Fanuc KAREL source: compact_preamble.KL

PROGRAM KB00046
%NOLOCKGROUP
%ENVIRONMENT FDEV
VAR
P1 : STRING[80];P2 : STRING[80];P3:BOOLEAN;P4:BOOLEAN;P5:INTEGER
BEGIN
P1='A'
P2='A'
P3=TRUE
P4=TRUE
P5=1
COPY_FILE(P1,P2,P3,P4,P5)
END KB00046
